// TIA Portal V21 export
// export: Created 2026-11-10T19:11:34.2261436Z, ExportSetting WithDefaults, DisplayName Totally Integrated Automation Portal, DisplayVersion V21 Update 3, DisplayName STEP 7 Professional, DisplayVersion V21 Update 3, DisplayName STEP 7 Safety, DisplayVersion V21, DisplayName Tech WebApplication, DisplayVersion V21, DisplayName WinCC Basic/Comfort/Advanced, DisplayVersion V21 Update 3, DisplayName WinCC Unified, DisplayVersion V21 Update 3
DATA_BLOCK "DB_TMAIL_C"   // DB14
// stored: AutoNumber true, DBAccessibleFromOPCUA true, DBAccessibleFromWebserver true, InstanceOfName TMAIL_C, OfSystemLibElement TMAIL_C, OfSystemLibVersion 6.1
"TMAIL_C"
   // VAR_INPUT
   //    REQ : Bool;
   //    TO_S : String[240];
   //    CC : String[240];
   //    SUBJECT : String[240];
   //    TEXT : String[240];
   //    ATTACHMENT : Variant;
   //    ATTACHMENT_NAME : String[50];
   //    MAIL_ADDR_PARAM : Variant;
   // END_VAR
   // VAR_OUTPUT
   //    DONE : Bool;
   //    BUSY : Bool;
   //    ERROR : Bool;
   //    STATUS : Word;
   // END_VAR
   // VAR
   //    SFB_STATUS : Word;
   //    PP : Int;
   //    Locked : Bool;
   //    RisingEdge : Bool;
   //    CpuInterface : Bool;
   //    WatchDogTime : Time;
   //    DiagCode : Word;
   //    MailObjectIndex : SInt;
   //    MailObjectCount : SInt;
   //    Byte_1 : Byte;
   //    UInt_1 : UInt;
   //    UDInt_1 : UDInt;
   //    UDInt_2 : UDInt;
   //    TMailDataHeader { S7_SetPoint := 'True'} : Array[1..7] of TMail_C_Header;
   //    T_MAIL { S7_SetPoint := 'True'} : T_MAIL;
   //    TCON { S7_SetPoint := 'True'} : TCON;
   //    TSEND { S7_SetPoint := 'True'} : TSEND;
   //    TRCV { S7_SetPoint := 'True'} : TRCV;
   //    TDISCON { S7_SetPoint := 'True'} : TDISCON;
   //    WatchDogTimer { S7_SetPoint := 'True'} : TON_TIME;
   // END_VAR
BEGIN
END_DATA_BLOCK
